Yaskawa INFORM job: LTEST.JBI

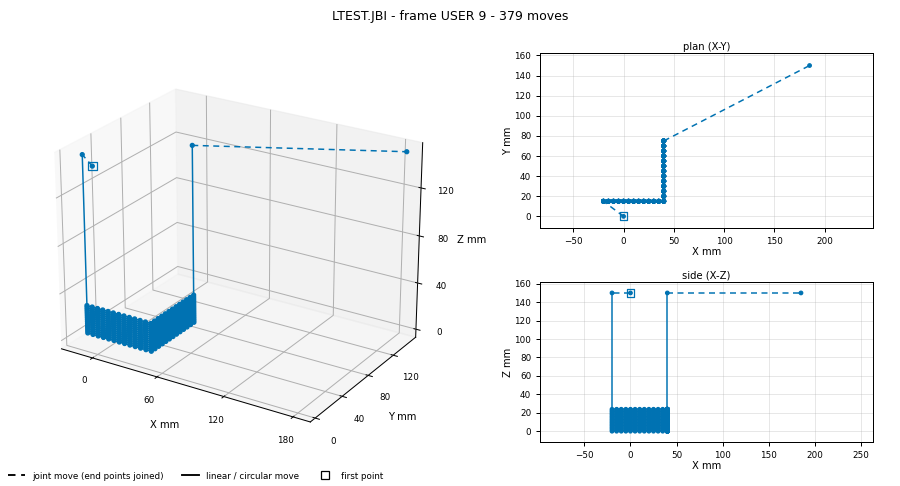
[picture p0: tool path of LTEST.JBI in frame USER 9, 379 of 379 moves have a stored position in this frame; points joined in program order, loops and branches not executed]
/JOB
//NAME LTEST
//POS
///NPOS 379,0,0,0,0,0
///USER 9
///TOOL 1
///POSTYPE USER
///RECTAN
///RCONF 1,0,0,0,0,0,0,0,0,0,0,0,0,0,0,0,0,0,0,0,0,0,0,0
C00000=0.000,0.000,150.000,0.0000,0.0000,-170.0000
C00001=-20.000,15.000,150.000,0.0000,0.0000,-170.0000
C00002=-20.000,15.000,0.000,0.0000,0.0000,-170.0000
C00003=-15.000,15.000,0.000,0.0000,0.0000,-170.0000
C00004=-10.000,15.000,0.000,0.0000,0.0000,-170.0000
C00005=-5.000,15.000,0.000,0.0000,0.0000,-170.0000
C00006=0.000,15.000,0.000,0.0000,0.0000,-170.0000
C00007=5.000,15.000,0.000,0.0000,0.0000,-170.0000
C00008=10.000,15.000,0.000,0.0000,0.0000,-170.0000
C00009=15.000,15.000,0.000,0.0000,0.0000,-170.0000
C00010=20.000,15.000,0.000,0.0000,0.0000,-170.0000
C00011=25.000,15.000,0.000,0.0000,0.0000,-170.0000
C00012=30.000,15.000,0.000,0.0000,0.0000,-170.0000
C00013=35.000,15.000,0.000,0.0000,0.0000,-170.0000
C00014=40.000,15.000,0.000,0.0000,0.0000,-170.0000
C00015=40.000,20.000,0.000,0.0000,0.0000,-170.0000
C00016=40.000,25.000,0.000,0.0000,0.0000,-170.0000
C00017=40.000,30.000,0.000,0.0000,0.0000,-170.0000
C00018=40.000,35.000,0.000,0.0000,0.0000,-170.0000
C00019=40.000,40.000,0.000,0.0000,0.0000,-170.0000
C00020=40.000,45.000,0.000,0.0000,0.0000,-170.0000
C00021=40.000,50.000,0.000,0.0000,0.0000,-170.0000
C00022=40.000,55.000,0.000,0.0000,0.0000,-170.0000
C00023=40.000,60.000,0.000,0.0000,0.0000,-170.0000
C00024=40.000,65.000,0.000,0.0000,0.0000,-170.0000
C00025=40.000,70.000,0.000,0.0000,0.0000,-170.0000
C00026=40.000,75.000,0.000,0.0000,0.0000,-170.0000
C00027=40.000,75.000,1.700,0.0000,0.0000,-170.0000
C00028=40.000,70.000,1.700,0.0000,0.0000,-170.0000
C00029=40.000,65.000,1.700,0.0000,0.0000,-170.0000
C00030=40.000,60.000,1.700,0.0000,0.0000,-170.0000
C00031=40.000,55.000,1.700,0.0000,0.0000,-170.0000
C00032=40.000,50.000,1.700,0.0000,0.0000,-170.0000
C00033=40.000,45.000,1.700,0.0000,0.0000,-170.0000
C00034=40.000,40.000,1.700,0.0000,0.0000,-170.0000
C00035=40.000,35.000,1.700,0.0000,0.0000,-170.0000
C00036=40.000,30.000,1.700,0.0000,0.0000,-170.0000
C00037=40.000,25.000,1.700,0.0000,0.0000,-170.0000
C00038=40.000,20.000,1.700,0.0000,0.0000,-170.0000
C00039=40.000,15.000,1.700,0.0000,0.0000,-170.0000
C00040=35.000,15.000,1.700,0.0000,0.0000,-170.0000
C00041=30.000,15.000,1.700,0.0000,0.0000,-170.0000
C00042=25.000,15.000,1.700,0.0000,0.0000,-170.0000
C00043=20.000,15.000,1.700,0.0000,0.0000,-170.0000
C00044=15.000,15.000,1.700,0.0000,0.0000,-170.0000
C00045=10.000,15.000,1.700,0.0000,0.0000,-170.0000
C00046=5.000,15.000,1.700,0.0000,0.0000,-170.0000
C00047=0.000,15.000,1.700,0.0000,0.0000,-170.0000
C00048=-5.000,15.000,1.700,0.0000,0.0000,-170.0000
C00049=-10.000,15.000,1.700,0.0000,0.0000,-170.0000
C00050=-15.000,15.000,1.700,0.0000,0.0000,-170.0000
C00051=-20.000,15.000,1.700,0.0000,0.0000,-170.0000
C00052=-20.000,15.000,3.400,0.0000,0.0000,-170.0000
C00053=-15.000,15.000,3.400,0.0000,0.0000,-170.0000
C00054=-10.000,15.000,3.400,0.0000,0.0000,-170.0000
C00055=-5.000,15.000,3.400,0.0000,0.0000,-170.0000
C00056=0.000,15.000,3.400,0.0000,0.0000,-170.0000
C00057=5.000,15.000,3.400,0.0000,0.0000,-170.0000
C00058=10.000,15.000,3.400,0.0000,0.0000,-170.0000
C00059=15.000,15.000,3.400,0.0000,0.0000,-170.0000
C00060=20.000,15.000,3.400,0.0000,0.0000,-170.0000
C00061=25.000,15.000,3.400,0.0000,0.0000,-170.0000
C00062=30.000,15.000,3.400,0.0000,0.0000,-170.0000
C00063=35.000,15.000,3.400,0.0000,0.0000,-170.0000
C00064=40.000,15.000,3.400,0.0000,0.0000,-170.0000
C00065=40.000,20.000,3.400,0.0000,0.0000,-170.0000
C00066=40.000,25.000,3.400,0.0000,0.0000,-170.0000
C00067=40.000,30.000,3.400,0.0000,0.0000,-170.0000
C00068=40.000,35.000,3.400,0.0000,0.0000,-170.0000
C00069=40.000,40.000,3.400,0.0000,0.0000,-170.0000
C00070=40.000,45.000,3.400,0.0000,0.0000,-170.0000
C00071=40.000,50.000,3.400,0.0000,0.0000,-170.0000
C00072=40.000,55.000,3.400,0.0000,0.0000,-170.0000
C00073=40.000,60.000,3.400,0.0000,0.0000,-170.0000
C00074=40.000,65.000,3.400,0.0000,0.0000,-170.0000
C00075=40.000,70.000,3.400,0.0000,0.0000,-170.0000
C00076=40.000,75.000,3.400,0.0000,0.0000,-170.0000
C00077=40.000,75.000,5.100,0.0000,0.0000,-170.0000
C00078=40.000,70.000,5.100,0.0000,0.0000,-170.0000
C00079=40.000,65.000,5.100,0.0000,0.0000,-170.0000
C00080=40.000,60.000,5.100,0.0000,0.0000,-170.0000
C00081=40.000,55.000,5.100,0.0000,0.0000,-170.0000
C00082=40.000,50.000,5.100,0.0000,0.0000,-170.0000
C00083=40.000,45.000,5.100,0.0000,0.0000,-170.0000
C00084=40.000,40.000,5.100,0.0000,0.0000,-170.0000
C00085=40.000,35.000,5.100,0.0000,0.0000,-170.0000
C00086=40.000,30.000,5.100,0.0000,0.0000,-170.0000
C00087=40.000,25.000,5.100,0.0000,0.0000,-170.0000
C00088=40.000,20.000,5.100,0.0000,0.0000,-170.0000
C00089=40.000,15.000,5.100,0.0000,0.0000,-170.0000
C00090=35.000,15.000,5.100,0.0000,0.0000,-170.0000
C00091=30.000,15.000,5.100,0.0000,0.0000,-170.0000
C00092=25.000,15.000,5.100,0.0000,0.0000,-170.0000
C00093=20.000,15.000,5.100,0.0000,0.0000,-170.0000
C00094=15.000,15.000,5.100,0.0000,0.0000,-170.0000
C00095=10.000,15.000,5.100,0.0000,0.0000,-170.0000
C00096=5.000,15.000,5.100,0.0000,0.0000,-170.0000
C00097=0.000,15.000,5.100,0.0000,0.0000,-170.0000
C00098=-5.000,15.000,5.100,0.0000,0.0000,-170.0000
C00099=-10.000,15.000,5.100,0.0000,0.0000,-170.0000
C00100=-15.000,15.000,5.100,0.0000,0.0000,-170.0000
C00101=-20.000,15.000,5.100,0.0000,0.0000,-170.0000
C00102=-20.000,15.000,6.800,0.0000,0.0000,-170.0000
C00103=-15.000,15.000,6.800,0.0000,0.0000,-170.0000
C00104=-10.000,15.000,6.800,0.0000,0.0000,-170.0000
C00105=-5.000,15.000,6.800,0.0000,0.0000,-170.0000
C00106=0.000,15.000,6.800,0.0000,0.0000,-170.0000
C00107=5.000,15.000,6.800,0.0000,0.0000,-170.0000
C00108=10.000,15.000,6.800,0.0000,0.0000,-170.0000
C00109=15.000,15.000,6.800,0.0000,0.0000,-170.0000
C00110=20.000,15.000,6.800,0.0000,0.0000,-170.0000
C00111=25.000,15.000,6.800,0.0000,0.0000,-170.0000
C00112=30.000,15.000,6.800,0.0000,0.0000,-170.0000
C00113=35.000,15.000,6.800,0.0000,0.0000,-170.0000
C00114=40.000,15.000,6.800,0.0000,0.0000,-170.0000
C00115=40.000,20.000,6.800,0.0000,0.0000,-170.0000
C00116=40.000,25.000,6.800,0.0000,0.0000,-170.0000
C00117=40.000,30.000,6.800,0.0000,0.0000,-170.0000
C00118=40.000,35.000,6.800,0.0000,0.0000,-170.0000
C00119=40.000,40.000,6.800,0.0000,0.0000,-170.0000
C00120=40.000,45.000,6.800,0.0000,0.0000,-170.0000
C00121=40.000,50.000,6.800,0.0000,0.0000,-170.0000
C00122=40.000,55.000,6.800,0.0000,0.0000,-170.0000
C00123=40.000,60.000,6.800,0.0000,0.0000,-170.0000
C00124=40.000,65.000,6.800,0.0000,0.0000,-170.0000
C00125=40.000,70.000,6.800,0.0000,0.0000,-170.0000
C00126=40.000,75.000,6.800,0.0000,0.0000,-170.0000
C00127=40.000,75.000,8.500,0.0000,0.0000,-170.0000
C00128=40.000,70.000,8.500,0.0000,0.0000,-170.0000
C00129=40.000,65.000,8.500,0.0000,0.0000,-170.0000
C00130=40.000,60.000,8.500,0.0000,0.0000,-170.0000
C00131=40.000,55.000,8.500,0.0000,0.0000,-170.0000
C00132=40.000,50.000,8.500,0.0000,0.0000,-170.0000
C00133=40.000,45.000,8.500,0.0000,0.0000,-170.0000
C00134=40.000,40.000,8.500,0.0000,0.0000,-170.0000
C00135=40.000,35.000,8.500,0.0000,0.0000,-170.0000
C00136=40.000,30.000,8.500,0.0000,0.0000,-170.0000
C00137=40.000,25.000,8.500,0.0000,0.0000,-170.0000
C00138=40.000,20.000,8.500,0.0000,0.0000,-170.0000
C00139=40.000,15.000,8.500,0.0000,0.0000,-170.0000
C00140=35.000,15.000,8.500,0.0000,0.0000,-170.0000
C00141=30.000,15.000,8.500,0.0000,0.0000,-170.0000
C00142=25.000,15.000,8.500,0.0000,0.0000,-170.0000
C00143=20.000,15.000,8.500,0.0000,0.0000,-170.0000
C00144=15.000,15.000,8.500,0.0000,0.0000,-170.0000
C00145=10.000,15.000,8.500,0.0000,0.0000,-170.0000
C00146=5.000,15.000,8.500,0.0000,0.0000,-170.0000
C00147=0.000,15.000,8.500,0.0000,0.0000,-170.0000
C00148=-5.000,15.000,8.500,0.0000,0.0000,-170.0000
C00149=-10.000,15.000,8.500,0.0000,0.0000,-170.0000
C00150=-15.000,15.000,8.500,0.0000,0.0000,-170.0000
C00151=-20.000,15.000,8.500,0.0000,0.0000,-170.0000
C00152=-20.000,15.000,10.200,0.0000,0.0000,-170.0000
C00153=-15.000,15.000,10.200,0.0000,0.0000,-170.0000
C00154=-10.000,15.000,10.200,0.0000,0.0000,-170.0000
C00155=-5.000,15.000,10.200,0.0000,0.0000,-170.0000
C00156=0.000,15.000,10.200,0.0000,0.0000,-170.0000
C00157=5.000,15.000,10.200,0.0000,0.0000,-170.0000
C00158=10.000,15.000,10.200,0.0000,0.0000,-170.0000
C00159=15.000,15.000,10.200,0.0000,0.0000,-170.0000
C00160=20.000,15.000,10.200,0.0000,0.0000,-170.0000
C00161=25.000,15.000,10.200,0.0000,0.0000,-170.0000
C00162=30.000,15.000,10.200,0.0000,0.0000,-170.0000
C00163=35.000,15.000,10.200,0.0000,0.0000,-170.0000
C00164=40.000,15.000,10.200,0.0000,0.0000,-170.0000
C00165=40.000,20.000,10.200,0.0000,0.0000,-170.0000
C00166=40.000,25.000,10.200,0.0000,0.0000,-170.0000
C00167=40.000,30.000,10.200,0.0000,0.0000,-170.0000
C00168=40.000,35.000,10.200,0.0000,0.0000,-170.0000
C00169=40.000,40.000,10.200,0.0000,0.0000,-170.0000
C00170=40.000,45.000,10.200,0.0000,0.0000,-170.0000
C00171=40.000,50.000,10.200,0.0000,0.0000,-170.0000
C00172=40.000,55.000,10.200,0.0000,0.0000,-170.0000
C00173=40.000,60.000,10.200,0.0000,0.0000,-170.0000
C00174=40.000,65.000,10.200,0.0000,0.0000,-170.0000
C00175=40.000,70.000,10.200,0.0000,0.0000,-170.0000
C00176=40.000,75.000,10.200,0.0000,0.0000,-170.0000
C00177=40.000,75.000,11.900,0.0000,0.0000,-170.0000
C00178=40.000,70.000,11.900,0.0000,0.0000,-170.0000
C00179=40.000,65.000,11.900,0.0000,0.0000,-170.0000
C00180=40.000,60.000,11.900,0.0000,0.0000,-170.0000
C00181=40.000,55.000,11.900,0.0000,0.0000,-170.0000
C00182=40.000,50.000,11.900,0.0000,0.0000,-170.0000
C00183=40.000,45.000,11.900,0.0000,0.0000,-170.0000
C00184=40.000,40.000,11.900,0.0000,0.0000,-170.0000
C00185=40.000,35.000,11.900,0.0000,0.0000,-170.0000
C00186=40.000,30.000,11.900,0.0000,0.0000,-170.0000
C00187=40.000,25.000,11.900,0.0000,0.0000,-170.0000
C00188=40.000,20.000,11.900,0.0000,0.0000,-170.0000
C00189=40.000,15.000,11.900,0.0000,0.0000,-170.0000
C00190=35.000,15.000,11.900,0.0000,0.0000,-170.0000
C00191=30.000,15.000,11.900,0.0000,0.0000,-170.0000
C00192=25.000,15.000,11.900,0.0000,0.0000,-170.0000
C00193=20.000,15.000,11.900,0.0000,0.0000,-170.0000
C00194=15.000,15.000,11.900,0.0000,0.0000,-170.0000
C00195=10.000,15.000,11.900,0.0000,0.0000,-170.0000
C00196=5.000,15.000,11.900,0.0000,0.0000,-170.0000
C00197=0.000,15.000,11.900,0.0000,0.0000,-170.0000
C00198=-5.000,15.000,11.900,0.0000,0.0000,-170.0000
C00199=-10.000,15.000,11.900,0.0000,0.0000,-170.0000
C00200=-15.000,15.000,11.900,0.0000,0.0000,-170.0000
C00201=-20.000,15.000,11.900,0.0000,0.0000,-170.0000
C00202=-20.000,15.000,13.600,0.0000,0.0000,-170.0000
C00203=-15.000,15.000,13.600,0.0000,0.0000,-170.0000
C00204=-10.000,15.000,13.600,0.0000,0.0000,-170.0000
C00205=-5.000,15.000,13.600,0.0000,0.0000,-170.0000
C00206=0.000,15.000,13.600,0.0000,0.0000,-170.0000
C00207=5.000,15.000,13.600,0.0000,0.0000,-170.0000
C00208=10.000,15.000,13.600,0.0000,0.0000,-170.0000
C00209=15.000,15.000,13.600,0.0000,0.0000,-170.0000
C00210=20.000,15.000,13.600,0.0000,0.0000,-170.0000
C00211=25.000,15.000,13.600,0.0000,0.0000,-170.0000
C00212=30.000,15.000,13.600,0.0000,0.0000,-170.0000
C00213=35.000,15.000,13.600,0.0000,0.0000,-170.0000
C00214=40.000,15.000,13.600,0.0000,0.0000,-170.0000
C00215=40.000,20.000,13.600,0.0000,0.0000,-170.0000
C00216=40.000,25.000,13.600,0.0000,0.0000,-170.0000
C00217=40.000,30.000,13.600,0.0000,0.0000,-170.0000
C00218=40.000,35.000,13.600,0.0000,0.0000,-170.0000
C00219=40.000,40.000,13.600,0.0000,0.0000,-170.0000
C00220=40.000,45.000,13.600,0.0000,0.0000,-170.0000
C00221=40.000,50.000,13.600,0.0000,0.0000,-170.0000
C00222=40.000,55.000,13.600,0.0000,0.0000,-170.0000
C00223=40.000,60.000,13.600,0.0000,0.0000,-170.0000
C00224=40.000,65.000,13.600,0.0000,0.0000,-170.0000
C00225=40.000,70.000,13.600,0.0000,0.0000,-170.0000
C00226=40.000,75.000,13.600,0.0000,0.0000,-170.0000
C00227=40.000,75.000,15.300,0.0000,0.0000,-170.0000
C00228=40.000,70.000,15.300,0.0000,0.0000,-170.0000
C00229=40.000,65.000,15.300,0.0000,0.0000,-170.0000
C00230=40.000,60.000,15.300,0.0000,0.0000,-170.0000
C00231=40.000,55.000,15.300,0.0000,0.0000,-170.0000
C00232=40.000,50.000,15.300,0.0000,0.0000,-170.0000
C00233=40.000,45.000,15.300,0.0000,0.0000,-170.0000
C00234=40.000,40.000,15.300,0.0000,0.0000,-170.0000
C00235=40.000,35.000,15.300,0.0000,0.0000,-170.0000
C00236=40.000,30.000,15.300,0.0000,0.0000,-170.0000
C00237=40.000,25.000,15.300,0.0000,0.0000,-170.0000
C00238=40.000,20.000,15.300,0.0000,0.0000,-170.0000
C00239=40.000,15.000,15.300,0.0000,0.0000,-170.0000
C00240=35.000,15.000,15.300,0.0000,0.0000,-170.0000
C00241=30.000,15.000,15.300,0.0000,0.0000,-170.0000
C00242=25.000,15.000,15.300,0.0000,0.0000,-170.0000
C00243=20.000,15.000,15.300,0.0000,0.0000,-170.0000
C00244=15.000,15.000,15.300,0.0000,0.0000,-170.0000
C00245=10.000,15.000,15.300,0.0000,0.0000,-170.0000
C00246=5.000,15.000,15.300,0.0000,0.0000,-170.0000
C00247=0.000,15.000,15.300,0.0000,0.0000,-170.0000
C00248=-5.000,15.000,15.300,0.0000,0.0000,-170.0000
C00249=-10.000,15.000,15.300,0.0000,0.0000,-170.0000
C00250=-15.000,15.000,15.300,0.0000,0.0000,-170.0000
C00251=-20.000,15.000,15.300,0.0000,0.0000,-170.0000
C00252=-20.000,15.000,17.000,0.0000,0.0000,-170.0000
C00253=-15.000,15.000,17.000,0.0000,0.0000,-170.0000
C00254=-10.000,15.000,17.000,0.0000,0.0000,-170.0000
C00255=-5.000,15.000,17.000,0.0000,0.0000,-170.0000
C00256=0.000,15.000,17.000,0.0000,0.0000,-170.0000
C00257=5.000,15.000,17.000,0.0000,0.0000,-170.0000
C00258=10.000,15.000,17.000,0.0000,0.0000,-170.0000
C00259=15.000,15.000,17.000,0.0000,0.0000,-170.0000
C00260=20.000,15.000,17.000,0.0000,0.0000,-170.0000
C00261=25.000,15.000,17.000,0.0000,0.0000,-170.0000
C00262=30.000,15.000,17.000,0.0000,0.0000,-170.0000
C00263=35.000,15.000,17.000,0.0000,0.0000,-170.0000
C00264=40.000,15.000,17.000,0.0000,0.0000,-170.0000
C00265=40.000,20.000,17.000,0.0000,0.0000,-170.0000
C00266=40.000,25.000,17.000,0.0000,0.0000,-170.0000
C00267=40.000,30.000,17.000,0.0000,0.0000,-170.0000
C00268=40.000,35.000,17.000,0.0000,0.0000,-170.0000
C00269=40.000,40.000,17.000,0.0000,0.0000,-170.0000
C00270=40.000,45.000,17.000,0.0000,0.0000,-170.0000
C00271=40.000,50.000,17.000,0.0000,0.0000,-170.0000
C00272=40.000,55.000,17.000,0.0000,0.0000,-170.0000
C00273=40.000,60.000,17.000,0.0000,0.0000,-170.0000
C00274=40.000,65.000,17.000,0.0000,0.0000,-170.0000
C00275=40.000,70.000,17.000,0.0000,0.0000,-170.0000
C00276=40.000,75.000,17.000,0.0000,0.0000,-170.0000
C00277=40.000,75.000,18.700,0.0000,0.0000,-170.0000
C00278=40.000,70.000,18.700,0.0000,0.0000,-170.0000
C00279=40.000,65.000,18.700,0.0000,0.0000,-170.0000
C00280=40.000,60.000,18.700,0.0000,0.0000,-170.0000
C00281=40.000,55.000,18.700,0.0000,0.0000,-170.0000
C00282=40.000,50.000,18.700,0.0000,0.0000,-170.0000
C00283=40.000,45.000,18.700,0.0000,0.0000,-170.0000
C00284=40.000,40.000,18.700,0.0000,0.0000,-170.0000
C00285=40.000,35.000,18.700,0.0000,0.0000,-170.0000
C00286=40.000,30.000,18.700,0.0000,0.0000,-170.0000
C00287=40.000,25.000,18.700,0.0000,0.0000,-170.0000
C00288=40.000,20.000,18.700,0.0000,0.0000,-170.0000
C00289=40.000,15.000,18.700,0.0000,0.0000,-170.0000
C00290=35.000,15.000,18.700,0.0000,0.0000,-170.0000
C00291=30.000,15.000,18.700,0.0000,0.0000,-170.0000
C00292=25.000,15.000,18.700,0.0000,0.0000,-170.0000
C00293=20.000,15.000,18.700,0.0000,0.0000,-170.0000
C00294=15.000,15.000,18.700,0.0000,0.0000,-170.0000
C00295=10.000,15.000,18.700,0.0000,0.0000,-170.0000
C00296=5.000,15.000,18.700,0.0000,0.0000,-170.0000
C00297=0.000,15.000,18.700,0.0000,0.0000,-170.0000
C00298=-5.000,15.000,18.700,0.0000,0.0000,-170.0000
C00299=-10.000,15.000,18.700,0.0000,0.0000,-170.0000
C00300=-15.000,15.000,18.700,0.0000,0.0000,-170.0000
C00301=-20.000,15.000,18.700,0.0000,0.0000,-170.0000
C00302=-20.000,15.000,20.400,0.0000,0.0000,-170.0000
C00303=-15.000,15.000,20.400,0.0000,0.0000,-170.0000
C00304=-10.000,15.000,20.400,0.0000,0.0000,-170.0000
C00305=-5.000,15.000,20.400,0.0000,0.0000,-170.0000
C00306=0.000,15.000,20.400,0.0000,0.0000,-170.0000
C00307=5.000,15.000,20.400,0.0000,0.0000,-170.0000
C00308=10.000,15.000,20.400,0.0000,0.0000,-170.0000
C00309=15.000,15.000,20.400,0.0000,0.0000,-170.0000
C00310=20.000,15.000,20.400,0.0000,0.0000,-170.0000
C00311=25.000,15.000,20.400,0.0000,0.0000,-170.0000
C00312=30.000,15.000,20.400,0.0000,0.0000,-170.0000
C00313=35.000,15.000,20.400,0.0000,0.0000,-170.0000
C00314=40.000,15.000,20.400,0.0000,0.0000,-170.0000
C00315=40.000,20.000,20.400,0.0000,0.0000,-170.0000
C00316=40.000,25.000,20.400,0.0000,0.0000,-170.0000
C00317=40.000,30.000,20.400,0.0000,0.0000,-170.0000
C00318=40.000,35.000,20.400,0.0000,0.0000,-170.0000
C00319=40.000,40.000,20.400,0.0000,0.0000,-170.0000
C00320=40.000,45.000,20.400,0.0000,0.0000,-170.0000
C00321=40.000,50.000,20.400,0.0000,0.0000,-170.0000
C00322=40.000,55.000,20.400,0.0000,0.0000,-170.0000
C00323=40.000,60.000,20.400,0.0000,0.0000,-170.0000
C00324=40.000,65.000,20.400,0.0000,0.0000,-170.0000
C00325=40.000,70.000,20.400,0.0000,0.0000,-170.0000
C00326=40.000,75.000,20.400,0.0000,0.0000,-170.0000
C00327=40.000,75.000,22.100,0.0000,0.0000,-170.0000
C00328=40.000,70.000,22.100,0.0000,0.0000,-170.0000
C00329=40.000,65.000,22.100,0.0000,0.0000,-170.0000
C00330=40.000,60.000,22.100,0.0000,0.0000,-170.0000
C00331=40.000,55.000,22.100,0.0000,0.0000,-170.0000
C00332=40.000,50.000,22.100,0.0000,0.0000,-170.0000
C00333=40.000,45.000,22.100,0.0000,0.0000,-170.0000
C00334=40.000,40.000,22.100,0.0000,0.0000,-170.0000
C00335=40.000,35.000,22.100,0.0000,0.0000,-170.0000
C00336=40.000,30.000,22.100,0.0000,0.0000,-170.0000
C00337=40.000,25.000,22.100,0.0000,0.0000,-170.0000
C00338=40.000,20.000,22.100,0.0000,0.0000,-170.0000
C00339=40.000,15.000,22.100,0.0000,0.0000,-170.0000
C00340=35.000,15.000,22.100,0.0000,0.0000,-170.0000
C00341=30.000,15.000,22.100,0.0000,0.0000,-170.0000
C00342=25.000,15.000,22.100,0.0000,0.0000,-170.0000
C00343=20.000,15.000,22.100,0.0000,0.0000,-170.0000
C00344=15.000,15.000,22.100,0.0000,0.0000,-170.0000
C00345=10.000,15.000,22.100,0.0000,0.0000,-170.0000
C00346=5.000,15.000,22.100,0.0000,0.0000,-170.0000
C00347=0.000,15.000,22.100,0.0000,0.0000,-170.0000
C00348=-5.000,15.000,22.100,0.0000,0.0000,-170.0000
C00349=-10.000,15.000,22.100,0.0000,0.0000,-170.0000
C00350=-15.000,15.000,22.100,0.0000,0.0000,-170.0000
C00351=-20.000,15.000,22.100,0.0000,0.0000,-170.0000
C00352=-20.000,15.000,23.800,0.0000,0.0000,-170.0000
C00353=-15.000,15.000,23.800,0.0000,0.0000,-170.0000
C00354=-10.000,15.000,23.800,0.0000,0.0000,-170.0000
C00355=-5.000,15.000,23.800,0.0000,0.0000,-170.0000
C00356=0.000,15.000,23.800,0.0000,0.0000,-170.0000
C00357=5.000,15.000,23.800,0.0000,0.0000,-170.0000
C00358=10.000,15.000,23.800,0.0000,0.0000,-170.0000
C00359=15.000,15.000,23.800,0.0000,0.0000,-170.0000
C00360=20.000,15.000,23.800,0.0000,0.0000,-170.0000
C00361=25.000,15.000,23.800,0.0000,0.0000,-170.0000
C00362=30.000,15.000,23.800,0.0000,0.0000,-170.0000
C00363=35.000,15.000,23.800,0.0000,0.0000,-170.0000
C00364=40.000,15.000,23.800,0.0000,0.0000,-170.0000
C00365=40.000,20.000,23.800,0.0000,0.0000,-170.0000
C00366=40.000,25.000,23.800,0.0000,0.0000,-170.0000
C00367=40.000,30.000,23.800,0.0000,0.0000,-170.0000
C00368=40.000,35.000,23.800,0.0000,0.0000,-170.0000
C00369=40.000,40.000,23.800,0.0000,0.0000,-170.0000
C00370=40.000,45.000,23.800,0.0000,0.0000,-170.0000
C00371=40.000,50.000,23.800,0.0000,0.0000,-170.0000
C00372=40.000,55.000,23.800,0.0000,0.0000,-170.0000
C00373=40.000,60.000,23.800,0.0000,0.0000,-170.0000
C00374=40.000,65.000,23.800,0.0000,0.0000,-170.0000
C00375=40.000,70.000,23.800,0.0000,0.0000,-170.0000
C00376=40.000,75.000,23.800,0.0000,0.0000,-170.0000
C00377=40.000,75.000,150.000,0.0000,0.0000,-170.0000
C00378=185.000,150.000,150.000,0.0000,0.0000,-170.0000
//INST
///DATE 2026/11/04 15:21
///ATTR SC,RW,RJ
////FRAME USER 9
///GROUP1 RB1
NOP
MOVJ C00000 VJ=0.78
MOVJ C00001 VJ=0.78
MOVL C00002 V=11.0 ACC=20 DEC=20
*LAG1
MACRO1 MJ#(0) ARGF1
ARCON
MOVL C00003 V=7.0 ACC=20 DEC=20
MOVL C00004 V=7.0 ACC=20 DEC=20
MOVL C00005 V=7.0 ACC=20 DEC=20
MOVL C00006 V=7.0 ACC=20 DEC=20
MOVL C00007 V=7.0 ACC=20 DEC=20
MOVL C00008 V=7.0 ACC=20 DEC=20
MOVL C00009 V=7.0 ACC=20 DEC=20
MOVL C00010 V=7.0 ACC=20 DEC=20
MOVL C00011 V=7.0 ACC=20 DEC=20
MOVL C00012 V=7.7 ACC=20 DEC=20
MOVL C00013 V=7.7 ACC=20 DEC=20
MOVL C00014 V=7.7 PL=1
MOVL C00015 V=7.7 ACC=20 DEC=20
MOVL C00016 V=7.7 ACC=20 DEC=20
MOVL C00017 V=7.0 ACC=20 DEC=20
MOVL C00018 V=7.0 ACC=20 DEC=20
MOVL C00019 V=7.0 ACC=20 DEC=20
MOVL C00020 V=7.0 ACC=20 DEC=20
MOVL C00021 V=7.0 ACC=20 DEC=20
MOVL C00022 V=7.0 ACC=20 DEC=20
MOVL C00023 V=7.0 ACC=20 DEC=20
MOVL C00024 V=7.0 ACC=20 DEC=20
MOVL C00025 V=7.0 ACC=20 DEC=20
MOVL C00026 V=7.0 ACC=20 DEC=20
ARCOF
TIMER T=30
MOVL C00027 V=11.0 ACC=20 DEC=20
*LAG2
MACRO1 MJ#(0) ARGF2
ARCON
MOVL C00028 V=7.0 ACC=20 DEC=20
MOVL C00029 V=7.0 ACC=20 DEC=20
MOVL C00030 V=7.0 ACC=20 DEC=20
MOVL C00031 V=7.0 ACC=20 DEC=20
MOVL C00032 V=7.0 ACC=20 DEC=20
MOVL C00033 V=7.0 ACC=20 DEC=20
MOVL C00034 V=7.0 ACC=20 DEC=20
MOVL C00035 V=7.0 ACC=20 DEC=20
MOVL C00036 V=7.0 ACC=20 DEC=20
MOVL C00037 V=7.7 ACC=20 DEC=20
MOVL C00038 V=7.7 ACC=20 DEC=20
MOVL C00039 V=7.7 PL=1
MOVL C00040 V=7.7 ACC=20 DEC=20
MOVL C00041 V=7.7 ACC=20 DEC=20
MOVL C00042 V=7.0 ACC=20 DEC=20
MOVL C00043 V=7.0 ACC=20 DEC=20
MOVL C00044 V=7.0 ACC=20 DEC=20
MOVL C00045 V=7.0 ACC=20 DEC=20
MOVL C00046 V=7.0 ACC=20 DEC=20
MOVL C00047 V=7.0 ACC=20 DEC=20
MOVL C00048 V=7.0 ACC=20 DEC=20
MOVL C00049 V=7.0 ACC=20 DEC=20
MOVL C00050 V=7.0 ACC=20 DEC=20
MOVL C00051 V=7.0 ACC=20 DEC=20
ARCOF
TIMER T=30
MOVL C00052 V=11.0 ACC=20 DEC=20
*LAG3
MACRO1 MJ#(0) ARGF2
ARCON
MOVL C00053 V=7.0 ACC=20 DEC=20
MOVL C00054 V=7.0 ACC=20 DEC=20
MOVL C00055 V=7.0 ACC=20 DEC=20
MOVL C00056 V=7.0 ACC=20 DEC=20
MOVL C00057 V=7.0 ACC=20 DEC=20
MOVL C00058 V=7.0 ACC=20 DEC=20
MOVL C00059 V=7.0 ACC=20 DEC=20
MOVL C00060 V=7.0 ACC=20 DEC=20
MOVL C00061 V=7.0 ACC=20 DEC=20
MOVL C00062 V=7.7 ACC=20 DEC=20
MOVL C00063 V=7.7 ACC=20 DEC=20
MOVL C00064 V=7.7 PL=1
MOVL C00065 V=7.7 ACC=20 DEC=20
MOVL C00066 V=7.7 ACC=20 DEC=20
MOVL C00067 V=7.0 ACC=20 DEC=20
MOVL C00068 V=7.0 ACC=20 DEC=20
MOVL C00069 V=7.0 ACC=20 DEC=20
MOVL C00070 V=7.0 ACC=20 DEC=20
MOVL C00071 V=7.0 ACC=20 DEC=20
MOVL C00072 V=7.0 ACC=20 DEC=20
MOVL C00073 V=7.0 ACC=20 DEC=20
MOVL C00074 V=7.0 ACC=20 DEC=20
MOVL C00075 V=7.0 ACC=20 DEC=20
MOVL C00076 V=7.0 ACC=20 DEC=20
ARCOF
TIMER T=30
MOVL C00077 V=11.0 ACC=20 DEC=20
*LAG4
MACRO1 MJ#(0) ARGF2
ARCON
MOVL C00078 V=7.0 ACC=20 DEC=20
MOVL C00079 V=7.0 ACC=20 DEC=20
MOVL C00080 V=7.0 ACC=20 DEC=20
MOVL C00081 V=7.0 ACC=20 DEC=20
MOVL C00082 V=7.0 ACC=20 DEC=20
MOVL C00083 V=7.0 ACC=20 DEC=20
MOVL C00084 V=7.0 ACC=20 DEC=20
MOVL C00085 V=7.0 ACC=20 DEC=20
MOVL C00086 V=7.0 ACC=20 DEC=20
MOVL C00087 V=7.7 ACC=20 DEC=20
MOVL C00088 V=7.7 ACC=20 DEC=20
MOVL C00089 V=7.7 PL=1
MOVL C00090 V=7.7 ACC=20 DEC=20
MOVL C00091 V=7.7 ACC=20 DEC=20
MOVL C00092 V=7.0 ACC=20 DEC=20
MOVL C00093 V=7.0 ACC=20 DEC=20
MOVL C00094 V=7.0 ACC=20 DEC=20
MOVL C00095 V=7.0 ACC=20 DEC=20
MOVL C00096 V=7.0 ACC=20 DEC=20
MOVL C00097 V=7.0 ACC=20 DEC=20
MOVL C00098 V=7.0 ACC=20 DEC=20
MOVL C00099 V=7.0 ACC=20 DEC=20
MOVL C00100 V=7.0 ACC=20 DEC=20
MOVL C00101 V=7.0 ACC=20 DEC=20
ARCOF
TIMER T=30
MOVL C00102 V=11.0 ACC=20 DEC=20
*LAG5
MACRO1 MJ#(0) ARGF2
ARCON
MOVL C00103 V=7.0 ACC=20 DEC=20
MOVL C00104 V=7.0 ACC=20 DEC=20
MOVL C00105 V=7.0 ACC=20 DEC=20
MOVL C00106 V=7.0 ACC=20 DEC=20
MOVL C00107 V=7.0 ACC=20 DEC=20
MOVL C00108 V=7.0 ACC=20 DEC=20
MOVL C00109 V=7.0 ACC=20 DEC=20
MOVL C00110 V=7.0 ACC=20 DEC=20
MOVL C00111 V=7.0 ACC=20 DEC=20
MOVL C00112 V=7.7 ACC=20 DEC=20
MOVL C00113 V=7.7 ACC=20 DEC=20
MOVL C00114 V=7.7 PL=1
MOVL C00115 V=7.7 ACC=20 DEC=20
MOVL C00116 V=7.7 ACC=20 DEC=20
MOVL C00117 V=7.0 ACC=20 DEC=20
MOVL C00118 V=7.0 ACC=20 DEC=20
MOVL C00119 V=7.0 ACC=20 DEC=20
MOVL C00120 V=7.0 ACC=20 DEC=20
MOVL C00121 V=7.0 ACC=20 DEC=20
MOVL C00122 V=7.0 ACC=20 DEC=20
MOVL C00123 V=7.0 ACC=20 DEC=20
MOVL C00124 V=7.0 ACC=20 DEC=20
MOVL C00125 V=7.0 ACC=20 DEC=20
MOVL C00126 V=7.0 ACC=20 DEC=20
ARCOF
TIMER T=30
MOVL C00127 V=11.0 ACC=20 DEC=20
*LAG6
MACRO1 MJ#(0) ARGF2
ARCON
MOVL C00128 V=7.0 ACC=20 DEC=20
MOVL C00129 V=7.0 ACC=20 DEC=20
MOVL C00130 V=7.0 ACC=20 DEC=20
MOVL C00131 V=7.0 ACC=20 DEC=20
MOVL C00132 V=7.0 ACC=20 DEC=20
MOVL C00133 V=7.0 ACC=20 DEC=20
MOVL C00134 V=7.0 ACC=20 DEC=20
MOVL C00135 V=7.0 ACC=20 DEC=20
MOVL C00136 V=7.0 ACC=20 DEC=20
MOVL C00137 V=7.7 ACC=20 DEC=20
MOVL C00138 V=7.7 ACC=20 DEC=20
MOVL C00139 V=7.7 PL=1
MOVL C00140 V=7.7 ACC=20 DEC=20
MOVL C00141 V=7.7 ACC=20 DEC=20
MOVL C00142 V=7.0 ACC=20 DEC=20
MOVL C00143 V=7.0 ACC=20 DEC=20
MOVL C00144 V=7.0 ACC=20 DEC=20
MOVL C00145 V=7.0 ACC=20 DEC=20
MOVL C00146 V=7.0 ACC=20 DEC=20
MOVL C00147 V=7.0 ACC=20 DEC=20
MOVL C00148 V=7.0 ACC=20 DEC=20
MOVL C00149 V=7.0 ACC=20 DEC=20
MOVL C00150 V=7.0 ACC=20 DEC=20
MOVL C00151 V=7.0 ACC=20 DEC=20
ARCOF
TIMER T=30
MOVL C00152 V=11.0 ACC=20 DEC=20
*LAG7
MACRO1 MJ#(0) ARGF2
ARCON
MOVL C00153 V=7.0 ACC=20 DEC=20
MOVL C00154 V=7.0 ACC=20 DEC=20
MOVL C00155 V=7.0 ACC=20 DEC=20
MOVL C00156 V=7.0 ACC=20 DEC=20
MOVL C00157 V=7.0 ACC=20 DEC=20
MOVL C00158 V=7.0 ACC=20 DEC=20
MOVL C00159 V=7.0 ACC=20 DEC=20
MOVL C00160 V=7.0 ACC=20 DEC=20
MOVL C00161 V=7.0 ACC=20 DEC=20
MOVL C00162 V=7.7 ACC=20 DEC=20
MOVL C00163 V=7.7 ACC=20 DEC=20
MOVL C00164 V=7.7 PL=1
MOVL C00165 V=7.7 ACC=20 DEC=20
MOVL C00166 V=7.7 ACC=20 DEC=20
MOVL C00167 V=7.0 ACC=20 DEC=20
MOVL C00168 V=7.0 ACC=20 DEC=20
MOVL C00169 V=7.0 ACC=20 DEC=20
MOVL C00170 V=7.0 ACC=20 DEC=20
MOVL C00171 V=7.0 ACC=20 DEC=20
MOVL C00172 V=7.0 ACC=20 DEC=20
MOVL C00173 V=7.0 ACC=20 DEC=20
MOVL C00174 V=7.0 ACC=20 DEC=20
MOVL C00175 V=7.0 ACC=20 DEC=20
MOVL C00176 V=7.0 ACC=20 DEC=20
ARCOF
TIMER T=30
MOVL C00177 V=11.0 ACC=20 DEC=20
*LAG8
MACRO1 MJ#(0) ARGF2
ARCON
MOVL C00178 V=7.0 ACC=20 DEC=20
MOVL C00179 V=7.0 ACC=20 DEC=20
MOVL C00180 V=7.0 ACC=20 DEC=20
MOVL C00181 V=7.0 ACC=20 DEC=20
MOVL C00182 V=7.0 ACC=20 DEC=20
MOVL C00183 V=7.0 ACC=20 DEC=20
MOVL C00184 V=7.0 ACC=20 DEC=20
MOVL C00185 V=7.0 ACC=20 DEC=20
MOVL C00186 V=7.0 ACC=20 DEC=20
MOVL C00187 V=7.7 ACC=20 DEC=20
MOVL C00188 V=7.7 ACC=20 DEC=20
MOVL C00189 V=7.7 PL=1
MOVL C00190 V=7.7 ACC=20 DEC=20
MOVL C00191 V=7.7 ACC=20 DEC=20
MOVL C00192 V=7.0 ACC=20 DEC=20
MOVL C00193 V=7.0 ACC=20 DEC=20
MOVL C00194 V=7.0 ACC=20 DEC=20
MOVL C00195 V=7.0 ACC=20 DEC=20
MOVL C00196 V=7.0 ACC=20 DEC=20
MOVL C00197 V=7.0 ACC=20 DEC=20
MOVL C00198 V=7.0 ACC=20 DEC=20
MOVL C00199 V=7.0 ACC=20 DEC=20
MOVL C00200 V=7.0 ACC=20 DEC=20
MOVL C00201 V=7.0 ACC=20 DEC=20
ARCOF
TIMER T=30
MOVL C00202 V=11.0 ACC=20 DEC=20
*LAG9
MACRO1 MJ#(0) ARGF2
ARCON
MOVL C00203 V=7.0 ACC=20 DEC=20
MOVL C00204 V=7.0 ACC=20 DEC=20
MOVL C00205 V=7.0 ACC=20 DEC=20
MOVL C00206 V=7.0 ACC=20 DEC=20
MOVL C00207 V=7.0 ACC=20 DEC=20
MOVL C00208 V=7.0 ACC=20 DEC=20
MOVL C00209 V=7.0 ACC=20 DEC=20
MOVL C00210 V=7.0 ACC=20 DEC=20
MOVL C00211 V=7.0 ACC=20 DEC=20
MOVL C00212 V=7.7 ACC=20 DEC=20
MOVL C00213 V=7.7 ACC=20 DEC=20
MOVL C00214 V=7.7 PL=1
MOVL C00215 V=7.7 ACC=20 DEC=20
MOVL C00216 V=7.7 ACC=20 DEC=20
MOVL C00217 V=7.0 ACC=20 DEC=20
MOVL C00218 V=7.0 ACC=20 DEC=20
MOVL C00219 V=7.0 ACC=20 DEC=20
MOVL C00220 V=7.0 ACC=20 DEC=20
MOVL C00221 V=7.0 ACC=20 DEC=20
MOVL C00222 V=7.0 ACC=20 DEC=20
MOVL C00223 V=7.0 ACC=20 DEC=20
MOVL C00224 V=7.0 ACC=20 DEC=20
MOVL C00225 V=7.0 ACC=20 DEC=20
MOVL C00226 V=7.0 ACC=20 DEC=20
ARCOF
TIMER T=30
MOVL C00227 V=11.0 ACC=20 DEC=20
*LAG10
MACRO1 MJ#(0) ARGF2
ARCON
MOVL C00228 V=7.0 ACC=20 DEC=20
MOVL C00229 V=7.0 ACC=20 DEC=20
MOVL C00230 V=7.0 ACC=20 DEC=20
MOVL C00231 V=7.0 ACC=20 DEC=20
MOVL C00232 V=7.0 ACC=20 DEC=20
MOVL C00233 V=7.0 ACC=20 DEC=20
MOVL C00234 V=7.0 ACC=20 DEC=20
MOVL C00235 V=7.0 ACC=20 DEC=20
MOVL C00236 V=7.0 ACC=20 DEC=20
MOVL C00237 V=7.7 ACC=20 DEC=20
MOVL C00238 V=7.7 ACC=20 DEC=20
MOVL C00239 V=7.7 PL=1
MOVL C00240 V=7.7 ACC=20 DEC=20
MOVL C00241 V=7.7 ACC=20 DEC=20
MOVL C00242 V=7.0 ACC=20 DEC=20
MOVL C00243 V=7.0 ACC=20 DEC=20
MOVL C00244 V=7.0 ACC=20 DEC=20
MOVL C00245 V=7.0 ACC=20 DEC=20
MOVL C00246 V=7.0 ACC=20 DEC=20
MOVL C00247 V=7.0 ACC=20 DEC=20
MOVL C00248 V=7.0 ACC=20 DEC=20
MOVL C00249 V=7.0 ACC=20 DEC=20
MOVL C00250 V=7.0 ACC=20 DEC=20
MOVL C00251 V=7.0 ACC=20 DEC=20
ARCOF
TIMER T=30
MOVL C00252 V=11.0 ACC=20 DEC=20
*LAG11
MACRO1 MJ#(0) ARGF2
ARCON
MOVL C00253 V=7.0 ACC=20 DEC=20
MOVL C00254 V=7.0 ACC=20 DEC=20
MOVL C00255 V=7.0 ACC=20 DEC=20
MOVL C00256 V=7.0 ACC=20 DEC=20
MOVL C00257 V=7.0 ACC=20 DEC=20
MOVL C00258 V=7.0 ACC=20 DEC=20
MOVL C00259 V=7.0 ACC=20 DEC=20
MOVL C00260 V=7.0 ACC=20 DEC=20
MOVL C00261 V=7.0 ACC=20 DEC=20
MOVL C00262 V=7.7 ACC=20 DEC=20
MOVL C00263 V=7.7 ACC=20 DEC=20
MOVL C00264 V=7.7 PL=1
MOVL C00265 V=7.7 ACC=20 DEC=20
MOVL C00266 V=7.7 ACC=20 DEC=20
MOVL C00267 V=7.0 ACC=20 DEC=20
MOVL C00268 V=7.0 ACC=20 DEC=20
MOVL C00269 V=7.0 ACC=20 DEC=20
MOVL C00270 V=7.0 ACC=20 DEC=20
MOVL C00271 V=7.0 ACC=20 DEC=20
MOVL C00272 V=7.0 ACC=20 DEC=20
MOVL C00273 V=7.0 ACC=20 DEC=20
MOVL C00274 V=7.0 ACC=20 DEC=20
MOVL C00275 V=7.0 ACC=20 DEC=20
MOVL C00276 V=7.0 ACC=20 DEC=20
ARCOF
TIMER T=30
MOVL C00277 V=11.0 ACC=20 DEC=20
*LAG12
MACRO1 MJ#(0) ARGF2
ARCON
MOVL C00278 V=7.0 ACC=20 DEC=20
MOVL C00279 V=7.0 ACC=20 DEC=20
MOVL C00280 V=7.0 ACC=20 DEC=20
MOVL C00281 V=7.0 ACC=20 DEC=20
MOVL C00282 V=7.0 ACC=20 DEC=20
MOVL C00283 V=7.0 ACC=20 DEC=20
MOVL C00284 V=7.0 ACC=20 DEC=20
MOVL C00285 V=7.0 ACC=20 DEC=20
MOVL C00286 V=7.0 ACC=20 DEC=20
MOVL C00287 V=7.7 ACC=20 DEC=20
MOVL C00288 V=7.7 ACC=20 DEC=20
MOVL C00289 V=7.7 PL=1
MOVL C00290 V=7.7 ACC=20 DEC=20
MOVL C00291 V=7.7 ACC=20 DEC=20
MOVL C00292 V=7.0 ACC=20 DEC=20
MOVL C00293 V=7.0 ACC=20 DEC=20
MOVL C00294 V=7.0 ACC=20 DEC=20
MOVL C00295 V=7.0 ACC=20 DEC=20
MOVL C00296 V=7.0 ACC=20 DEC=20
MOVL C00297 V=7.0 ACC=20 DEC=20
MOVL C00298 V=7.0 ACC=20 DEC=20
MOVL C00299 V=7.0 ACC=20 DEC=20
MOVL C00300 V=7.0 ACC=20 DEC=20
MOVL C00301 V=7.0 ACC=20 DEC=20
ARCOF
TIMER T=30
MOVL C00302 V=11.0 ACC=20 DEC=20
*LAG13
MACRO1 MJ#(0) ARGF2
ARCON
MOVL C00303 V=7.0 ACC=20 DEC=20
MOVL C00304 V=7.0 ACC=20 DEC=20
MOVL C00305 V=7.0 ACC=20 DEC=20
MOVL C00306 V=7.0 ACC=20 DEC=20
MOVL C00307 V=7.0 ACC=20 DEC=20
MOVL C00308 V=7.0 ACC=20 DEC=20
MOVL C00309 V=7.0 ACC=20 DEC=20
MOVL C00310 V=7.0 ACC=20 DEC=20
MOVL C00311 V=7.0 ACC=20 DEC=20
MOVL C00312 V=7.7 ACC=20 DEC=20
MOVL C00313 V=7.7 ACC=20 DEC=20
MOVL C00314 V=7.7 PL=1
MOVL C00315 V=7.7 ACC=20 DEC=20
MOVL C00316 V=7.7 ACC=20 DEC=20
MOVL C00317 V=7.0 ACC=20 DEC=20
MOVL C00318 V=7.0 ACC=20 DEC=20
MOVL C00319 V=7.0 ACC=20 DEC=20
MOVL C00320 V=7.0 ACC=20 DEC=20
MOVL C00321 V=7.0 ACC=20 DEC=20
MOVL C00322 V=7.0 ACC=20 DEC=20
MOVL C00323 V=7.0 ACC=20 DEC=20
MOVL C00324 V=7.0 ACC=20 DEC=20
MOVL C00325 V=7.0 ACC=20 DEC=20
MOVL C00326 V=7.0 ACC=20 DEC=20
ARCOF
TIMER T=30
MOVL C00327 V=11.0 ACC=20 DEC=20
*LAG14
MACRO1 MJ#(0) ARGF2
ARCON
MOVL C00328 V=7.0 ACC=20 DEC=20
MOVL C00329 V=7.0 ACC=20 DEC=20
MOVL C00330 V=7.0 ACC=20 DEC=20
MOVL C00331 V=7.0 ACC=20 DEC=20
MOVL C00332 V=7.0 ACC=20 DEC=20
MOVL C00333 V=7.0 ACC=20 DEC=20
MOVL C00334 V=7.0 ACC=20 DEC=20
MOVL C00335 V=7.0 ACC=20 DEC=20
MOVL C00336 V=7.0 ACC=20 DEC=20
MOVL C00337 V=7.7 ACC=20 DEC=20
MOVL C00338 V=7.7 ACC=20 DEC=20
MOVL C00339 V=7.7 PL=1
MOVL C00340 V=7.7 ACC=20 DEC=20
MOVL C00341 V=7.7 ACC=20 DEC=20
MOVL C00342 V=7.0 ACC=20 DEC=20
MOVL C00343 V=7.0 ACC=20 DEC=20
MOVL C00344 V=7.0 ACC=20 DEC=20
MOVL C00345 V=7.0 ACC=20 DEC=20
MOVL C00346 V=7.0 ACC=20 DEC=20
MOVL C00347 V=7.0 ACC=20 DEC=20
MOVL C00348 V=7.0 ACC=20 DEC=20
MOVL C00349 V=7.0 ACC=20 DEC=20
MOVL C00350 V=7.0 ACC=20 DEC=20
MOVL C00351 V=7.0 ACC=20 DEC=20
ARCOF
TIMER T=30
MOVL C00352 V=11.0 ACC=20 DEC=20
*LAG15
MACRO1 MJ#(0) ARGF2
ARCON
MOVL C00353 V=7.0 ACC=20 DEC=20
MOVL C00354 V=7.0 ACC=20 DEC=20
MOVL C00355 V=7.0 ACC=20 DEC=20
MOVL C00356 V=7.0 ACC=20 DEC=20
MOVL C00357 V=7.0 ACC=20 DEC=20
MOVL C00358 V=7.0 ACC=20 DEC=20
MOVL C00359 V=7.0 ACC=20 DEC=20
MOVL C00360 V=7.0 ACC=20 DEC=20
MOVL C00361 V=7.0 ACC=20 DEC=20
MOVL C00362 V=7.7 ACC=20 DEC=20
MOVL C00363 V=7.7 ACC=20 DEC=20
MOVL C00364 V=7.7 PL=1
MOVL C00365 V=7.7 ACC=20 DEC=20
MOVL C00366 V=7.7 ACC=20 DEC=20
MOVL C00367 V=7.0 ACC=20 DEC=20
MOVL C00368 V=7.0 ACC=20 DEC=20
MOVL C00369 V=7.0 ACC=20 DEC=20
MOVL C00370 V=7.0 ACC=20 DEC=20
MOVL C00371 V=7.0 ACC=20 DEC=20
MOVL C00372 V=7.0 ACC=20 DEC=20
MOVL C00373 V=7.0 ACC=20 DEC=20
MOVL C00374 V=7.0 ACC=20 DEC=20
MOVL C00375 V=7.0 ACC=20 DEC=20
MOVL C00376 V=7.0 ACC=20 DEC=20
ARCOF
TIMER T=30
MOVL C00377 V=11.0 ACC=20 DEC=20
MOVJ C00378 VJ=0.78
END
